(* IEC 61131-3 sources: Trarbach/resolucao/entrega/plc_corrigido, 1 file *)

(* ---- Prova2_corrigido.st ---- *)
(* Prova2_corrigido.st: Prova2.st com derivada filtrada. Unicas alteracoes: variaveis VP_F e kf_VP e o bloco
   marcado CORRECAO 1/2 antes do bloco DERIVATIVE. Validado so em simulacao (plc_sim.py), nao na bancada. *)
PROGRAM PI_D
  VAR
    SC : UINT;
  END_VAR
  VAR
    VP AT %IW0 : UINT;
    SP AT %QW0 : UINT;
    SO AT %QW1 : UINT := 6800;
  END_VAR
  VAR
    SO_AUX : UINT;
  END_VAR
  VAR
    MF AT %QX0.0 : BOOL := 0;
  END_VAR
  VAR
    VP_PERC : REAL;
    SP_PERC : REAL;
    SO_PERC : REAL;
    SC_PERC : REAL;
    SO_MAIS_P_INT_DER_PERC : REAL;
    ERRO_PERC : REAL;
    Kp_ERRO_PERC : REAL;
    Ki_ERRO_PERC : REAL;
    Ki_intgrERRO_PERC : REAL;
    Kd_VP_PERC : REAL;
    Kd_derVP_PERC : REAL;
    M_ACAO : REAL := 1.0;
    kp : REAL := 3.523;
    ki : REAL := 0.03872;
    kd : REAL := 39.16;
    STOP_INTGR : BOOL := 0;
    INTEGRAL_SEM_CI : INTEGRAL;
    DERIVADA : DERIVATIVE;
    SP_ant : REAL := 0.0;
    var_SP : REAL := 0.0;
    alfa : REAL := 1.0;
    FF2GL : REAL := 0.0;
    VP_F : REAL := 0.0;
    kf_VP : REAL := 0.017699;
    MMRY : UINT := 0;
    _TMP_SUB89_OUT : REAL;
    _TMP_MUL90_OUT : REAL;
    _TMP_SEL103_OUT : REAL;
    _TMP_ABS139_OUT : REAL;
    _TMP_LT137_OUT : BOOL;
    _TMP_SEL140_OUT : REAL;
    _TMP_MUL63_OUT : REAL;
    _TMP_MUL99_OUT : REAL;
    _TMP_SEL41_OUT : REAL;
    _TMP_MUL24_OUT : REAL;
    _TMP_MUL113_OUT : REAL;
    _TMP_SEL1_OUT : REAL;
    _TMP_MUL109_OUT : REAL;
    _TMP_ADD97_OUT : REAL;
    _TMP_ADD66_OUT : REAL;
    _TMP_SUB162_OUT : REAL;
    _TMP_GE34_OUT : BOOL;
    _TMP_LE4_OUT : BOOL;
    _TMP_OR44_OUT : BOOL;
    _TMP_LIMIT27_OUT : REAL;
    _TMP_SEL18_OUT : UINT;
    _TMP_SEL50_OUT : UINT;
    _TMP_SEL26_OUT : UINT;
    _TMP_UINT_TO_REAL68_OUT : REAL;
    _TMP_MUL69_OUT : REAL;
    _TMP_UINT_TO_REAL71_OUT : REAL;
    _TMP_MUL72_OUT : REAL;
    _TMP_MUL78_OUT : REAL;
    _TMP_REAL_TO_UINT77_OUT : UINT;
    _TMP_UINT_TO_REAL74_OUT : REAL;
    _TMP_MUL75_OUT : REAL;
    _TMP_NE148_OUT : BOOL;
    _TMP_SUB149_OUT : REAL;
    _TMP_SEL150_OUT : REAL;
    _TMP_SEL171_OUT : REAL;
    _TMP_SEL151_OUT : REAL;
    _TMP_AND169_OUT : BOOL;
    _TMP_SUB178_OUT : REAL;
    _TMP_MUL157_OUT : REAL;
    _TMP_SEL165_OUT : REAL;
    _TMP_ADD167_OUT : REAL;
    _TMP_SEL173_OUT : REAL;
    _TMP_MUL180_OUT : REAL;
    _TMP_REAL_TO_UINT182_OUT : UINT;
  END_VAR

  _TMP_SUB89_OUT := SUB(SP_PERC, VP_PERC);
  _TMP_MUL90_OUT := MUL(_TMP_SUB89_OUT, M_ACAO);
  _TMP_SEL103_OUT := SEL(MF, 0.0, _TMP_MUL90_OUT);
  _TMP_ABS139_OUT := ABS(_TMP_SEL103_OUT);
  _TMP_LT137_OUT := LT(_TMP_ABS139_OUT, 0.09);
  _TMP_SEL140_OUT := SEL(_TMP_LT137_OUT, _TMP_SEL103_OUT, 0.0);
  ERRO_PERC := _TMP_SEL140_OUT;
  _TMP_MUL63_OUT := MUL(ERRO_PERC, ki);
  Ki_ERRO_PERC := _TMP_MUL63_OUT;
  _TMP_MUL99_OUT := MUL(ERRO_PERC, kp);
  Kp_ERRO_PERC := _TMP_MUL99_OUT;
  _TMP_SEL41_OUT := SEL(STOP_INTGR, Ki_ERRO_PERC, 0.0);
  INTEGRAL_SEM_CI(RUN := TRUE, R1 := NOT(MF), XIN := _TMP_SEL41_OUT, X0 := 0.0, CYCLE := T#500ms);
  _TMP_MUL24_OUT := MUL(INTEGRAL_SEM_CI.XOUT, 0.04);
  Ki_intgrERRO_PERC := _TMP_MUL24_OUT;
  (* CORRECAO 1: passa-baixa de 1a ordem na VP antes da derivada (kf_VP = Ts/(tauf+Ts) = 0.02/(1.11+0.02); tauf = mu*Td = 1.11 s; Ts = 20 ms).
     Em manual VP_F acompanha a VP. *)
  IF NOT MF THEN
    VP_F := VP_PERC;
  ELSE
    VP_F := VP_F + kf_VP * (VP_PERC - VP_F);
  END_IF;
  (* CORRECAO 2: sem SEL(MF, 0.0, ...): a derivada fica 'armada' tambem em manual,
     eliminando o pulso de 3 scans ao fechar a malha. *)
  _TMP_MUL113_OUT := MUL(-1.0, VP_F, kd, M_ACAO);
  _TMP_SEL1_OUT := _TMP_MUL113_OUT;
  Kd_VP_PERC := _TMP_SEL1_OUT;
  DERIVADA(RUN := TRUE, XIN := Kd_VP_PERC, CYCLE := T#500ms);
  _TMP_MUL109_OUT := MUL(DERIVADA.XOUT, 25.0);
  Kd_derVP_PERC := _TMP_MUL109_OUT;
  _TMP_ADD97_OUT := ADD(Kp_ERRO_PERC, Ki_intgrERRO_PERC, Kd_derVP_PERC);
  _TMP_ADD66_OUT := ADD(_TMP_ADD97_OUT, SO_PERC);
  _TMP_SUB162_OUT := SUB(_TMP_ADD66_OUT, FF2GL);
  SO_MAIS_P_INT_DER_PERC := _TMP_SUB162_OUT;
  _TMP_GE34_OUT := GE(SO_MAIS_P_INT_DER_PERC, 100.0);
  _TMP_LE4_OUT := LE(SO_MAIS_P_INT_DER_PERC, 10.0);
  _TMP_OR44_OUT := OR(_TMP_GE34_OUT, _TMP_LE4_OUT);
  STOP_INTGR := _TMP_OR44_OUT;
  _TMP_LIMIT27_OUT := LIMIT(10.0, SO_MAIS_P_INT_DER_PERC, 100.0);
  SC_PERC := _TMP_LIMIT27_OUT;
  _TMP_SEL18_OUT := SEL(MF, SO, SO_AUX);
  SO_AUX := _TMP_SEL18_OUT;
  _TMP_SEL50_OUT := SEL(MF, VP, SP);
  SP := _TMP_SEL50_OUT;
  _TMP_SEL26_OUT := SEL(MF, SO, SC);
  SO := _TMP_SEL26_OUT;
  _TMP_UINT_TO_REAL68_OUT := UINT_TO_REAL(VP);
  _TMP_MUL69_OUT := MUL(_TMP_UINT_TO_REAL68_OUT, 0.001525);
  VP_PERC := _TMP_MUL69_OUT;
  _TMP_UINT_TO_REAL71_OUT := UINT_TO_REAL(SP);
  _TMP_MUL72_OUT := MUL(_TMP_UINT_TO_REAL71_OUT, 0.001525);
  SP_PERC := _TMP_MUL72_OUT;
  _TMP_MUL78_OUT := MUL(SC_PERC, 655.35);
  _TMP_REAL_TO_UINT77_OUT := REAL_TO_UINT(_TMP_MUL78_OUT);
  SC := _TMP_REAL_TO_UINT77_OUT;
  _TMP_UINT_TO_REAL74_OUT := UINT_TO_REAL(SO_AUX);
  _TMP_MUL75_OUT := MUL(_TMP_UINT_TO_REAL74_OUT, 0.001525);
  SO_PERC := _TMP_MUL75_OUT;
  _TMP_NE148_OUT := NE(SP_PERC, SP_ant);
  _TMP_SUB149_OUT := SUB(SP_PERC, SP_ant);
  _TMP_SEL150_OUT := SEL(_TMP_NE148_OUT, var_SP, _TMP_SUB149_OUT);
  _TMP_SEL171_OUT := SEL(MF, 0.0, _TMP_SEL150_OUT);
  var_SP := _TMP_SEL171_OUT;
  _TMP_SEL151_OUT := SEL(_TMP_NE148_OUT, SP_ant, SP_PERC);
  SP_ant := _TMP_SEL151_OUT;
  _TMP_AND169_OUT := AND(_TMP_NE148_OUT, MF);
  _TMP_SUB178_OUT := SUB(1.0, alfa);
  _TMP_MUL157_OUT := MUL(kp, _TMP_SUB178_OUT, var_SP);
  _TMP_SEL165_OUT := SEL(_TMP_AND169_OUT, 0.0, _TMP_MUL157_OUT);
  _TMP_ADD167_OUT := ADD(_TMP_SEL165_OUT, FF2GL);
  _TMP_SEL173_OUT := SEL(MF, 0.0, _TMP_ADD167_OUT);
  FF2GL := _TMP_SEL173_OUT;
  _TMP_MUL180_OUT := MUL(alfa, 25700.0);
  _TMP_REAL_TO_UINT182_OUT := REAL_TO_UINT(_TMP_MUL180_OUT);
  MMRY := _TMP_REAL_TO_UINT182_OUT;
END_PROGRAM

CONFIGURATION Config0

  RESOURCE Res0 ON PLC
    TASK task0(INTERVAL := T#20ms,PRIORITY := 0);
    PROGRAM instance0 WITH task0 : PI_D;
  END_RESOURCE
END_CONFIGURATION
